(* IEC 61131-3 sources: iecf/tools/bench, 28 files *)

(* ---- fbcalls.st ---- *)
(* iecf's benchmark (docs/testing/performance.md): 10 instances of a FUNCTION_BLOCK and a FUNCTION called 50 times a cycle, a CTU.
   Standard IEC 61131-3, for both compilers: tools/bench/run.sh. *)
FUNCTION_BLOCK Filter
  VAR_INPUT x : DINT; k : DINT; END_VAR
  VAR_OUTPUT y : DINT; END_VAR
  VAR state : DINT; n : DINT; END_VAR
  state := state + (x - state) / k;
  n := n + 1;
  y := state + n MOD 7;
END_FUNCTION_BLOCK
FUNCTION Mix : DINT
  VAR_INPUT a : DINT; b : DINT; END_VAR
  Mix := (a * 3 + b) MOD 100003;
END_FUNCTION
PROGRAM main
  VAR f1 : Filter; f2 : Filter; f3 : Filter; f4 : Filter; f5 : Filter; f6 : Filter; f7 : Filter; f8 : Filter; f9 : Filter; f10 : Filter; c : CTU; i : INT; rep : INT; acc : DINT; END_VAR
  VAR o1 AT %QD0 : DINT; o2 AT %QW4 : INT; END_VAR
  FOR rep := 1 TO 50 DO
    FOR i := 1 TO 10 DO
      f1(x := acc + 1, k := 4);
      acc := Mix(a := acc, b := f1.y);
      f2(x := acc + 2, k := 4);
      acc := Mix(a := acc, b := f2.y);
      f3(x := acc + 3, k := 4);
      acc := Mix(a := acc, b := f3.y);
      f4(x := acc + 4, k := 4);
      acc := Mix(a := acc, b := f4.y);
      f5(x := acc + 5, k := 4);
      acc := Mix(a := acc, b := f5.y);
      f6(x := acc + 6, k := 4);
      acc := Mix(a := acc, b := f6.y);
      f7(x := acc + 7, k := 4);
      acc := Mix(a := acc, b := f7.y);
      f8(x := acc + 8, k := 4);
      acc := Mix(a := acc, b := f8.y);
      f9(x := acc + 9, k := 4);
      acc := Mix(a := acc, b := f9.y);
      f10(x := acc + 10, k := 4);
      acc := Mix(a := acc, b := f10.y);
    END_FOR;
    c(CU := NOT c.CU, PV := 30000);
  END_FOR;
  IF c.Q THEN c(R := TRUE); c(R := FALSE); END_IF;
  o1 := acc;
  o2 := c.CV;
END_PROGRAM
CONFIGURATION cf
  RESOURCE r ON x
    TASK tk(INTERVAL := T#10ms, PRIORITY := 1);
    PROGRAM p WITH tk : main;
  END_RESOURCE
END_CONFIGURATION

(* ---- m_fbcall.st ---- *)
(* iecf's benchmark (docs/testing/performance.md): a FUNCTION_BLOCK call.
   Standard IEC 61131-3, for both compilers: tools/bench/run.sh. *)
FUNCTION_BLOCK Acc
  VAR_INPUT x : DINT; k : DINT; END_VAR
  VAR_OUTPUT y : DINT; END_VAR
  y := (y + x * k) MOD 100000;
END_FUNCTION_BLOCK
PROGRAM main
  VAR i : DINT; f : Acc; n : DINT; END_VAR
  VAR o1 AT %QD0 : DINT; END_VAR
  FOR i := 1 TO 20000 DO
    f(x := i MOD 9, k := 2); n := f.y;
  END_FOR;
  o1 := n;
END_PROGRAM
CONFIGURATION cf
  RESOURCE r ON x
    TASK tk(INTERVAL := T#10ms, PRIORITY := 1);
    PROGRAM p WITH tk : main;
  END_RESOURCE
END_CONFIGURATION

(* ---- oo.st ---- *)
(* iecf's benchmark (docs/testing/performance.md): CODESYS's object
   orientation, iecf alone (--extension codesys): set `mode` to 0 for a
   method of an instance, 1 through an interface, 2 through a REFERENCE
   TO, 3 through a POINTER TO, 4 a property read through an interface. *)
INTERFACE ICounter
  METHOD Bump : DINT
    VAR_INPUT amount : DINT; END_VAR
  END_METHOD
  PROPERTY Value : DINT
  GET
  END_GET
  END_PROPERTY
END_INTERFACE
FUNCTION_BLOCK Base IMPLEMENTS ICounter
  VAR n : DINT; END_VAR
  METHOD PUBLIC Bump : DINT
    VAR_INPUT amount : DINT; END_VAR
    n := (n + amount) MOD 100003;
    Bump := n;
  END_METHOD
  PROPERTY PUBLIC Value : DINT
  GET
    Value := n;
  END_GET
  END_PROPERTY
END_FUNCTION_BLOCK
FUNCTION_BLOCK Derived EXTENDS Base
  METHOD PUBLIC Bump : DINT
    VAR_INPUT amount : DINT; END_VAR
    n := (n + amount * 2) MOD 100003;
    Bump := n;
  END_METHOD
END_FUNCTION_BLOCK
PROGRAM main
  VAR i : DINT; b : Base; d : Derived; c : ICounter; r : REFERENCE TO Base; p : POINTER TO Base;
      acc : DINT; mode : DINT; END_VAR
  VAR o1 AT %QD0 : DINT; END_VAR
  r REF= d;
  p := ADR(b);
  FOR i := 1 TO 20000 DO
    CASE mode OF
      0: acc := acc + b.Bump(amount := i MOD 7);
      1: c := d; acc := acc + c.Bump(amount := i MOD 7);
      2: acc := acc + r.Bump(amount := i MOD 7);
      3: acc := acc + p^.Bump(amount := i MOD 7);
      4: c := b; acc := acc + c.Value;
    END_CASE;
    acc := acc MOD 1000003;
  END_FOR;
  o1 := acc;
END_PROGRAM
CONFIGURATION cf
  RESOURCE r ON x
    TASK tk(INTERVAL := T#10ms, PRIORITY := 1);
    PROGRAM p WITH tk : main;
  END_RESOURCE
END_CONFIGURATION

(* ---- sfc.st ---- *)
(* iecf's benchmark (docs/testing/performance.md): 40 instances of a FUNCTION_BLOCK whose body is a four-step SFC chart of N actions.
   Standard IEC 61131-3, for both compilers: tools/bench/run.sh. *)
FUNCTION_BLOCK Machine
  VAR_INPUT seed : DINT; END_VAR
  VAR_OUTPUT work : DINT; cycles : DINT; END_VAR
  VAR n : DINT; acc : DINT; END_VAR
  INITIAL_STEP idle : start(N); END_STEP
  TRANSITION FROM idle TO fill := n >= 2; END_TRANSITION
  STEP fill : filling(N); END_STEP
  TRANSITION FROM fill TO heat := n >= 5; END_TRANSITION
  STEP heat : heating(N); END_STEP
  TRANSITION FROM heat TO drain := n >= 9; END_TRANSITION
  STEP drain : draining(N); END_STEP
  TRANSITION FROM drain TO idle := n >= 12; END_TRANSITION
  ACTION start :
    n := n + 1;
    acc := (acc * 7 + seed) MOD 100003;
    work := acc;
  END_ACTION
  ACTION filling :
    n := n + 1;
    acc := (acc + seed * 3) MOD 100003;
    work := acc;
  END_ACTION
  ACTION heating :
    n := n + 1;
    acc := (acc * 3 + 11) MOD 100003;
    work := acc;
  END_ACTION
  ACTION draining :
    n := n + 1;
    IF n >= 12 THEN n := 0; cycles := cycles + 1; END_IF;
    acc := (acc + 5) MOD 100003;
    work := acc;
  END_ACTION
END_FUNCTION_BLOCK
PROGRAM main
  VAR m1 : Machine; m2 : Machine; m3 : Machine; m4 : Machine; m5 : Machine; m6 : Machine; m7 : Machine; m8 : Machine; m9 : Machine; m10 : Machine; m11 : Machine; m12 : Machine; m13 : Machine; m14 : Machine; m15 : Machine; m16 : Machine; m17 : Machine; m18 : Machine; m19 : Machine; m20 : Machine; m21 : Machine; m22 : Machine; m23 : Machine; m24 : Machine; m25 : Machine; m26 : Machine; m27 : Machine; m28 : Machine; m29 : Machine; m30 : Machine; m31 : Machine; m32 : Machine; m33 : Machine; m34 : Machine; m35 : Machine; m36 : Machine; m37 : Machine; m38 : Machine; m39 : Machine; m40 : Machine; total : DINT; c : DINT; END_VAR
  VAR o1 AT %QD0 : DINT; o2 AT %QD4 : DINT; END_VAR
  total := 0; c := 0;
  m1(seed := 1); total := (total + m1.work) MOD 1000003; c := c + m1.cycles;
  m2(seed := 2); total := (total + m2.work) MOD 1000003; c := c + m2.cycles;
  m3(seed := 3); total := (total + m3.work) MOD 1000003; c := c + m3.cycles;
  m4(seed := 4); total := (total + m4.work) MOD 1000003; c := c + m4.cycles;
  m5(seed := 5); total := (total + m5.work) MOD 1000003; c := c + m5.cycles;
  m6(seed := 6); total := (total + m6.work) MOD 1000003; c := c + m6.cycles;
  m7(seed := 7); total := (total + m7.work) MOD 1000003; c := c + m7.cycles;
  m8(seed := 8); total := (total + m8.work) MOD 1000003; c := c + m8.cycles;
  m9(seed := 9); total := (total + m9.work) MOD 1000003; c := c + m9.cycles;
  m10(seed := 10); total := (total + m10.work) MOD 1000003; c := c + m10.cycles;
  m11(seed := 11); total := (total + m11.work) MOD 1000003; c := c + m11.cycles;
  m12(seed := 12); total := (total + m12.work) MOD 1000003; c := c + m12.cycles;
  m13(seed := 13); total := (total + m13.work) MOD 1000003; c := c + m13.cycles;
  m14(seed := 14); total := (total + m14.work) MOD 1000003; c := c + m14.cycles;
  m15(seed := 15); total := (total + m15.work) MOD 1000003; c := c + m15.cycles;
  m16(seed := 16); total := (total + m16.work) MOD 1000003; c := c + m16.cycles;
  m17(seed := 17); total := (total + m17.work) MOD 1000003; c := c + m17.cycles;
  m18(seed := 18); total := (total + m18.work) MOD 1000003; c := c + m18.cycles;
  m19(seed := 19); total := (total + m19.work) MOD 1000003; c := c + m19.cycles;
  m20(seed := 20); total := (total + m20.work) MOD 1000003; c := c + m20.cycles;
  m21(seed := 21); total := (total + m21.work) MOD 1000003; c := c + m21.cycles;
  m22(seed := 22); total := (total + m22.work) MOD 1000003; c := c + m22.cycles;
  m23(seed := 23); total := (total + m23.work) MOD 1000003; c := c + m23.cycles;
  m24(seed := 24); total := (total + m24.work) MOD 1000003; c := c + m24.cycles;
  m25(seed := 25); total := (total + m25.work) MOD 1000003; c := c + m25.cycles;
  m26(seed := 26); total := (total + m26.work) MOD 1000003; c := c + m26.cycles;
  m27(seed := 27); total := (total + m27.work) MOD 1000003; c := c + m27.cycles;
  m28(seed := 28); total := (total + m28.work) MOD 1000003; c := c + m28.cycles;
  m29(seed := 29); total := (total + m29.work) MOD 1000003; c := c + m29.cycles;
  m30(seed := 30); total := (total + m30.work) MOD 1000003; c := c + m30.cycles;
  m31(seed := 31); total := (total + m31.work) MOD 1000003; c := c + m31.cycles;
  m32(seed := 32); total := (total + m32.work) MOD 1000003; c := c + m32.cycles;
  m33(seed := 33); total := (total + m33.work) MOD 1000003; c := c + m33.cycles;
  m34(seed := 34); total := (total + m34.work) MOD 1000003; c := c + m34.cycles;
  m35(seed := 35); total := (total + m35.work) MOD 1000003; c := c + m35.cycles;
  m36(seed := 36); total := (total + m36.work) MOD 1000003; c := c + m36.cycles;
  m37(seed := 37); total := (total + m37.work) MOD 1000003; c := c + m37.cycles;
  m38(seed := 38); total := (total + m38.work) MOD 1000003; c := c + m38.cycles;
  m39(seed := 39); total := (total + m39.work) MOD 1000003; c := c + m39.cycles;
  m40(seed := 40); total := (total + m40.work) MOD 1000003; c := c + m40.cycles;
  o1 := total;
  o2 := c;
END_PROGRAM
CONFIGURATION cf
  RESOURCE r ON x
    TASK tk(INTERVAL := T#10ms, PRIORITY := 1);
    PROGRAM p WITH tk : main;
  END_RESOURCE
END_CONFIGURATION

(* ---- arith.st ---- *)
(* iecf's benchmark (docs/testing/performance.md): integer and LREAL arithmetic in a loop: DINT products and MOD, ROL and XOR of a DWORD, SQRT.
   Standard IEC 61131-3, for both compilers: tools/bench/run.sh. *)
PROGRAM main
  VAR i : DINT; acc : DINT; w : DWORD := 16#1234567; x : LREAL; END_VAR
  VAR o1 AT %QD0 : DINT; o2 AT %QD4 : DINT; o3 AT %QD8 : DWORD; END_VAR
  FOR i := 1 TO 20000 DO
    acc := (acc * 31 + i) MOD 1000003;
    w := ROL(w, 3) XOR DINT_TO_DWORD(i);
    x := x + SQRT(DINT_TO_LREAL(i)) * 0.5;
  END_FOR;
  IF x > 1.0E9 THEN x := 0.0; END_IF;
  o1 := acc;
  o2 := LREAL_TO_DINT(x);
  o3 := w;
END_PROGRAM
CONFIGURATION cf
  RESOURCE r ON x
    TASK tk(INTERVAL := T#10ms, PRIORITY := 1);
    PROGRAM p WITH tk : main;
  END_RESOURCE
END_CONFIGURATION

(* ---- m_bool.st ---- *)
(* iecf's benchmark (docs/testing/performance.md): BOOL logic and IF.
   Standard IEC 61131-3, for both compilers: tools/bench/run.sh. *)

PROGRAM main
  VAR i : DINT; b : BOOL; c : BOOL; n : DINT; END_VAR
  VAR o1 AT %QD0 : DINT; END_VAR
  FOR i := 1 TO 20000 DO
    b := (i MOD 3 = 0) XOR c; IF b AND NOT c THEN n := n + 1; END_IF; c := b OR (i MOD 5 = 1);
  END_FOR;
  o1 := n;
END_PROGRAM
CONFIGURATION cf
  RESOURCE r ON x
    TASK tk(INTERVAL := T#10ms, PRIORITY := 1);
    PROGRAM p WITH tk : main;
  END_RESOURCE
END_CONFIGURATION

(* ---- m_case.st ---- *)
(* iecf's benchmark (docs/testing/performance.md): CASE with lists and ranges.
   Standard IEC 61131-3, for both compilers: tools/bench/run.sh. *)

PROGRAM main
  VAR i : DINT; n : DINT; END_VAR
  VAR o1 AT %QD0 : DINT; END_VAR
  FOR i := 1 TO 20000 DO
    CASE i MOD 8 OF 0: n := n + 1; 1, 2: n := n + 2; 3..5: n := n - 1; ELSE n := n + 3; END_CASE;
  END_FOR;
  o1 := n;
END_PROGRAM
CONFIGURATION cf
  RESOURCE r ON x
    TASK tk(INTERVAL := T#10ms, PRIORITY := 1);
    PROGRAM p WITH tk : main;
  END_RESOURCE
END_CONFIGURATION

(* ---- m_empty.st ---- *)
(* iecf's benchmark (docs/testing/performance.md): one statement: the cost of a cycle itself.
   Standard IEC 61131-3, for both compilers: tools/bench/run.sh. *)
PROGRAM main
  VAR n : DINT; END_VAR
  VAR o1 AT %QD0 : DINT; END_VAR
  n := n + 1;
  o1 := n;
END_PROGRAM
CONFIGURATION cf
  RESOURCE r ON x
    TASK tk(INTERVAL := T#10ms, PRIORITY := 1);
    PROGRAM p WITH tk : main;
  END_RESOURCE
END_CONFIGURATION

(* ---- m_fcall.st ---- *)
(* iecf's benchmark (docs/testing/performance.md): a FUNCTION call.
   Standard IEC 61131-3, for both compilers: tools/bench/run.sh. *)
FUNCTION Add3 : DINT
  VAR_INPUT a : DINT; b : DINT; c : DINT; END_VAR
  Add3 := a + b + c;
END_FUNCTION
PROGRAM main
  VAR i : DINT; n : DINT; END_VAR
  VAR o1 AT %QD0 : DINT; END_VAR
  FOR i := 1 TO 20000 DO
    n := Add3(a := n, b := i, c := 1) MOD 100000;
  END_FOR;
  o1 := n;
END_PROGRAM
CONFIGURATION cf
  RESOURCE r ON x
    TASK tk(INTERVAL := T#10ms, PRIORITY := 1);
    PROGRAM p WITH tk : main;
  END_RESOURCE
END_CONFIGURATION

(* ---- m_iadd.st ---- *)
(* iecf's benchmark (docs/testing/performance.md): a DINT sum.
   Standard IEC 61131-3, for both compilers: tools/bench/run.sh. *)

PROGRAM main
  VAR i : DINT; acc : DINT; END_VAR
  VAR o1 AT %QD0 : DINT; END_VAR
  FOR i := 1 TO 20000 DO
    acc := acc + i MOD 7;
  END_FOR;
  o1 := acc;
END_PROGRAM
CONFIGURATION cf
  RESOURCE r ON x
    TASK tk(INTERVAL := T#10ms, PRIORITY := 1);
    PROGRAM p WITH tk : main;
  END_RESOURCE
END_CONFIGURATION

(* ---- m_iarr.st ---- *)
(* iecf's benchmark (docs/testing/performance.md): a DINT array element updated.
   Standard IEC 61131-3, for both compilers: tools/bench/run.sh. *)

PROGRAM main
  VAR i : DINT; a : ARRAY[0..63] OF DINT; k : DINT; END_VAR
  VAR o1 AT %QD0 : DINT; END_VAR
  FOR i := 1 TO 20000 DO
    k := i MOD 64; a[k] := a[k] + i MOD 5;
  END_FOR;
  o1 := a[3];
END_PROGRAM
CONFIGURATION cf
  RESOURCE r ON x
    TASK tk(INTERVAL := T#10ms, PRIORITY := 1);
    PROGRAM p WITH tk : main;
  END_RESOURCE
END_CONFIGURATION

(* ---- m_imul.st ---- *)
(* iecf's benchmark (docs/testing/performance.md): a DINT product and MOD.
   Standard IEC 61131-3, for both compilers: tools/bench/run.sh. *)

PROGRAM main
  VAR i : DINT; acc : DINT := 1; END_VAR
  VAR o1 AT %QD0 : DINT; END_VAR
  FOR i := 1 TO 20000 DO
    acc := (acc * 3 + i) MOD 65521;
  END_FOR;
  o1 := acc;
END_PROGRAM
CONFIGURATION cf
  RESOURCE r ON x
    TASK tk(INTERVAL := T#10ms, PRIORITY := 1);
    PROGRAM p WITH tk : main;
  END_RESOURCE
END_CONFIGURATION

(* ---- m_lradd.st ---- *)
(* iecf's benchmark (docs/testing/performance.md): an LREAL sum.
   Standard IEC 61131-3, for both compilers: tools/bench/run.sh. *)

PROGRAM main
  VAR i : DINT; x : LREAL; s : LREAL; END_VAR
  VAR o1 AT %QD0 : DINT; END_VAR
  FOR i := 1 TO 20000 DO
    x := DINT_TO_LREAL(i); s := s + x;
  END_FOR;
  o1 := LREAL_TO_DINT(s / 1000.0);
END_PROGRAM
CONFIGURATION cf
  RESOURCE r ON x
    TASK tk(INTERVAL := T#10ms, PRIORITY := 1);
    PROGRAM p WITH tk : main;
  END_RESOURCE
END_CONFIGURATION

(* ---- m_str.st ---- *)
(* iecf's benchmark (docs/testing/performance.md): CONCAT and LEN.
   Standard IEC 61131-3, for both compilers: tools/bench/run.sh. *)

PROGRAM main
  VAR i : DINT; s : STRING; n : DINT; END_VAR
  VAR o1 AT %QD0 : DINT; END_VAR
  FOR i := 1 TO 20000 DO
    s := CONCAT('ab', 'cd'); n := n + LEN(s);
  END_FOR;
  o1 := n;
END_PROGRAM
CONFIGURATION cf
  RESOURCE r ON x
    TASK tk(INTERVAL := T#10ms, PRIORITY := 1);
    PROGRAM p WITH tk : main;
  END_RESOURCE
END_CONFIGURATION

(* ---- m_struct.st ---- *)
(* iecf's benchmark (docs/testing/performance.md): a structure assigned field by field and copied.
   Standard IEC 61131-3, for both compilers: tools/bench/run.sh. *)
TYPE Pt : STRUCT x : DINT; y : DINT; END_STRUCT; END_TYPE
PROGRAM main
  VAR i : DINT; p : Pt; q : Pt; n : DINT; END_VAR
  VAR o1 AT %QD0 : DINT; END_VAR
  FOR i := 1 TO 20000 DO
    p.x := i; p.y := i MOD 9; q := p; n := (n + q.x + q.y) MOD 100000;
  END_FOR;
  o1 := n;
END_PROGRAM
CONFIGURATION cf
  RESOURCE r ON x
    TASK tk(INTERVAL := T#10ms, PRIORITY := 1);
    PROGRAM p WITH tk : main;
  END_RESOURCE
END_CONFIGURATION

(* ---- m_ton.st ---- *)
(* iecf's benchmark (docs/testing/performance.md): a TON called.
   Standard IEC 61131-3, for both compilers: tools/bench/run.sh. *)

PROGRAM main
  VAR i : DINT; t : TON; n : DINT; END_VAR
  VAR o1 AT %QD0 : DINT; END_VAR
  FOR i := 1 TO 20000 DO
    t(IN := i MOD 2 = 0, PT := T#5ms); IF t.Q THEN n := n + 1; END_IF;
  END_FOR;
  o1 := n;
END_PROGRAM
CONFIGURATION cf
  RESOURCE r ON x
    TASK tk(INTERVAL := T#10ms, PRIORITY := 1);
    PROGRAM p WITH tk : main;
  END_RESOURCE
END_CONFIGURATION

(* ---- m_while.st ---- *)
(* iecf's benchmark (docs/testing/performance.md): a WHILE loop.
   Standard IEC 61131-3, for both compilers: tools/bench/run.sh. *)

PROGRAM main
  VAR i : DINT; j : DINT; n : DINT; END_VAR
  VAR o1 AT %QD0 : DINT; END_VAR
  FOR i := 1 TO 20000 DO
    j := i MOD 8; WHILE j > 0 DO n := n + j; j := j - 1; END_WHILE;
  END_FOR;
  o1 := n;
END_PROGRAM
CONFIGURATION cf
  RESOURCE r ON x
    TASK tk(INTERVAL := T#10ms, PRIORITY := 1);
    PROGRAM p WITH tk : main;
  END_RESOURCE
END_CONFIGURATION

(* ---- r_arr.st ---- *)
(* iecf's benchmark (docs/testing/performance.md): a REAL array element updated through a computed index.
   Standard IEC 61131-3, for both compilers: tools/bench/run.sh. *)
PROGRAM main
  VAR i : DINT; k : INT; x : LREAL; s : LREAL; r : REAL; arr : ARRAY[1..64] OF REAL; END_VAR
  VAR o1 AT %QD0 : DINT; o2 AT %QD4 : DINT; o3 AT %QD8 : DINT; END_VAR
  FOR i := 1 TO 5000 DO
    x := DINT_TO_LREAL(i) * 0.001;
    k := DINT_TO_INT(i MOD 64) + 1; arr[k] := arr[k] * 0.5 + r / 1000.0; r := r + 0.25;
  END_FOR;
  IF s > 1.0E9 THEN s := 0.0; END_IF;
  o1 := LREAL_TO_DINT(s);
  o2 := REAL_TO_DINT(r);
  o3 := REAL_TO_DINT(arr[7] * 100.0);
END_PROGRAM
CONFIGURATION cf
  RESOURCE r ON x
    TASK tk(INTERVAL := T#10ms, PRIORITY := 1);
    PROGRAM p WITH tk : main;
  END_RESOURCE
END_CONFIGURATION

(* ---- r_conv.st ---- *)
(* iecf's benchmark (docs/testing/performance.md): one statement each: an LREAL product of a DINT, an LREAL sum.
   Standard IEC 61131-3, for both compilers: tools/bench/run.sh. *)
PROGRAM main
  VAR i : DINT; k : INT; x : LREAL; s : LREAL; r : REAL; arr : ARRAY[1..64] OF REAL; END_VAR
  VAR o1 AT %QD0 : DINT; o2 AT %QD4 : DINT; o3 AT %QD8 : DINT; END_VAR
  FOR i := 1 TO 5000 DO
    x := DINT_TO_LREAL(i) * 0.001;
    s := s + x;
  END_FOR;
  IF s > 1.0E9 THEN s := 0.0; END_IF;
  o1 := LREAL_TO_DINT(s);
  o2 := REAL_TO_DINT(r);
  o3 := REAL_TO_DINT(arr[7] * 100.0);
END_PROGRAM
CONFIGURATION cf
  RESOURCE r ON x
    TASK tk(INTERVAL := T#10ms, PRIORITY := 1);
    PROGRAM p WITH tk : main;
  END_RESOURCE
END_CONFIGURATION

(* ---- r_explog.st ---- *)
(* iecf's benchmark (docs/testing/performance.md): EXP of a negated variable plus LN.
   Standard IEC 61131-3, for both compilers: tools/bench/run.sh. *)
PROGRAM main
  VAR i : DINT; k : INT; x : LREAL; s : LREAL; r : REAL; arr : ARRAY[1..64] OF REAL; END_VAR
  VAR o1 AT %QD0 : DINT; o2 AT %QD4 : DINT; o3 AT %QD8 : DINT; END_VAR
  FOR i := 1 TO 5000 DO
    x := DINT_TO_LREAL(i) * 0.001;
    s := s + EXP(-x) + LN(1.0 + x);
  END_FOR;
  IF s > 1.0E9 THEN s := 0.0; END_IF;
  o1 := LREAL_TO_DINT(s);
  o2 := REAL_TO_DINT(r);
  o3 := REAL_TO_DINT(arr[7] * 100.0);
END_PROGRAM
CONFIGURATION cf
  RESOURCE r ON x
    TASK tk(INTERVAL := T#10ms, PRIORITY := 1);
    PROGRAM p WITH tk : main;
  END_RESOURCE
END_CONFIGURATION

(* ---- r_real.st ---- *)
(* iecf's benchmark (docs/testing/performance.md): a REAL product plus an LREAL converted.
   Standard IEC 61131-3, for both compilers: tools/bench/run.sh. *)
PROGRAM main
  VAR i : DINT; k : INT; x : LREAL; s : LREAL; r : REAL; arr : ARRAY[1..64] OF REAL; END_VAR
  VAR o1 AT %QD0 : DINT; o2 AT %QD4 : DINT; o3 AT %QD8 : DINT; END_VAR
  FOR i := 1 TO 5000 DO
    x := DINT_TO_LREAL(i) * 0.001;
    r := r * 0.999 + LREAL_TO_REAL(x);
  END_FOR;
  IF s > 1.0E9 THEN s := 0.0; END_IF;
  o1 := LREAL_TO_DINT(s);
  o2 := REAL_TO_DINT(r);
  o3 := REAL_TO_DINT(arr[7] * 100.0);
END_PROGRAM
CONFIGURATION cf
  RESOURCE r ON x
    TASK tk(INTERVAL := T#10ms, PRIORITY := 1);
    PROGRAM p WITH tk : main;
  END_RESOURCE
END_CONFIGURATION

(* ---- r_sincos.st ---- *)
(* iecf's benchmark (docs/testing/performance.md): SIN times COS.
   Standard IEC 61131-3, for both compilers: tools/bench/run.sh. *)
PROGRAM main
  VAR i : DINT; k : INT; x : LREAL; s : LREAL; r : REAL; arr : ARRAY[1..64] OF REAL; END_VAR
  VAR o1 AT %QD0 : DINT; o2 AT %QD4 : DINT; o3 AT %QD8 : DINT; END_VAR
  FOR i := 1 TO 5000 DO
    x := DINT_TO_LREAL(i) * 0.001;
    s := s + SIN(x) * COS(x);
  END_FOR;
  IF s > 1.0E9 THEN s := 0.0; END_IF;
  o1 := LREAL_TO_DINT(s);
  o2 := REAL_TO_DINT(r);
  o3 := REAL_TO_DINT(arr[7] * 100.0);
END_PROGRAM
CONFIGURATION cf
  RESOURCE r ON x
    TASK tk(INTERVAL := T#10ms, PRIORITY := 1);
    PROGRAM p WITH tk : main;
  END_RESOURCE
END_CONFIGURATION

(* ---- r_sqrtdiv.st ---- *)
(* iecf's benchmark (docs/testing/performance.md): SQRT divided by a sum.
   Standard IEC 61131-3, for both compilers: tools/bench/run.sh. *)
PROGRAM main
  VAR i : DINT; k : INT; x : LREAL; s : LREAL; r : REAL; arr : ARRAY[1..64] OF REAL; END_VAR
  VAR o1 AT %QD0 : DINT; o2 AT %QD4 : DINT; o3 AT %QD8 : DINT; END_VAR
  FOR i := 1 TO 5000 DO
    x := DINT_TO_LREAL(i) * 0.001;
    s := s + SQRT(x) / (1.0 + x * x);
  END_FOR;
  IF s > 1.0E9 THEN s := 0.0; END_IF;
  o1 := LREAL_TO_DINT(s);
  o2 := REAL_TO_DINT(r);
  o3 := REAL_TO_DINT(arr[7] * 100.0);
END_PROGRAM
CONFIGURATION cf
  RESOURCE r ON x
    TASK tk(INTERVAL := T#10ms, PRIORITY := 1);
    PROGRAM p WITH tk : main;
  END_RESOURCE
END_CONFIGURATION

(* ---- reals.st ---- *)
(* iecf's benchmark (docs/testing/performance.md): LREAL SIN, COS, EXP, LN, SQRT and a division, a REAL array, 5000 times a cycle.
   Standard IEC 61131-3, for both compilers: tools/bench/run.sh. *)
PROGRAM main
  VAR i : DINT; k : INT; x : LREAL; s : LREAL; r : REAL; arr : ARRAY[1..64] OF REAL; END_VAR
  VAR o1 AT %QD0 : DINT; o2 AT %QD4 : DINT; o3 AT %QD8 : DINT; END_VAR
  FOR i := 1 TO 5000 DO
    x := DINT_TO_LREAL(i) * 0.001;
    s := s + SIN(x) * COS(x) + EXP(-x) + LN(1.0 + x) + SQRT(x) / (1.0 + x * x);
    r := r * 0.999 + LREAL_TO_REAL(x);
    k := DINT_TO_INT(i MOD 64) + 1;
    arr[k] := arr[k] * 0.5 + r / 1000.0;
  END_FOR;
  IF s > 1.0E9 THEN s := 0.0; END_IF;
  o1 := LREAL_TO_DINT(s);
  o2 := REAL_TO_DINT(r);
  o3 := REAL_TO_DINT(arr[7] * 100.0);
END_PROGRAM
CONFIGURATION cf
  RESOURCE r ON x
    TASK tk(INTERVAL := T#10ms, PRIORITY := 1);
    PROGRAM p WITH tk : main;
  END_RESOURCE
END_CONFIGURATION

(* ---- realsf.st ---- *)
(* iecf's benchmark (docs/testing/performance.md): `reals` in REAL - SIN, COS, EXP, LN, SQRT and a division, a REAL array, 5000 times a cycle.
   Standard IEC 61131-3, for both compilers: tools/bench/run.sh. *)
PROGRAM main
  VAR i : DINT; k : INT; x : REAL; s : REAL; r : REAL; arr : ARRAY[1..64] OF REAL; END_VAR
  VAR o1 AT %QD0 : DINT; o2 AT %QD4 : DINT; o3 AT %QD8 : DINT; END_VAR
  FOR i := 1 TO 5000 DO
    x := DINT_TO_REAL(i) * 0.001;
    s := s + SIN(x) * COS(x) + EXP(-x) + LN(1.0 + x) + SQRT(x) / (1.0 + x * x);
    r := r * 0.999 + x;
    k := DINT_TO_INT(i MOD 64) + 1;
    arr[k] := arr[k] * 0.5 + r / 1000.0;
  END_FOR;
  IF s > 1.0E9 THEN s := 0.0; END_IF;
  o1 := REAL_TO_DINT(s);
  o2 := REAL_TO_DINT(r);
  o3 := REAL_TO_DINT(arr[7] * 100.0);
END_PROGRAM
CONFIGURATION cf
  RESOURCE r ON x
    TASK tk(INTERVAL := T#10ms, PRIORITY := 1);
    PROGRAM p WITH tk : main;
  END_RESOURCE
END_CONFIGURATION

(* ---- sort.st ---- *)
(* iecf's benchmark (docs/testing/performance.md): an insertion sort of 300 DINTs, filled by a linear congruential generator.
   Standard IEC 61131-3, for both compilers: tools/bench/run.sh. *)
PROGRAM main
  VAR a : ARRAY[1..300] OF DINT; i : INT; j : INT; k : DINT; seed : DINT := 7; sum : DINT; END_VAR
  VAR o1 AT %QD0 : DINT; o2 AT %QD4 : DINT; END_VAR
  FOR i := 1 TO 300 DO
    seed := (seed * 1103 + 12345) MOD 65536;
    a[i] := seed;
  END_FOR;
  FOR i := 2 TO 300 DO
    k := a[i];
    j := i - 1;
    WHILE j >= 1 DO
      IF a[j] <= k THEN EXIT; END_IF;
      a[j + 1] := a[j];
      j := j - 1;
    END_WHILE;
    a[j + 1] := k;
  END_FOR;
  sum := 0;
  FOR i := 1 TO 300 DO sum := (sum + a[i] * INT_TO_DINT(i)) MOD 1000003; END_FOR;
  o1 := sum;
  o2 := a[150];
END_PROGRAM
CONFIGURATION cf
  RESOURCE r ON x
    TASK tk(INTERVAL := T#10ms, PRIORITY := 1);
    PROGRAM p WITH tk : main;
  END_RESOURCE
END_CONFIGURATION

(* ---- strings.st ---- *)
(* iecf's benchmark (docs/testing/performance.md): CONCAT, LEFT, RIGHT, LEN, FIND, INT_TO_STRING and STRING_TO_INT, 1000 times a cycle.
   Standard IEC 61131-3, for both compilers: tools/bench/run.sh. *)
PROGRAM main
  VAR i : INT; s : STRING; t : STRING := 'pump-station-'; n : DINT; END_VAR
  VAR o1 AT %QD0 : DINT; END_VAR
  FOR i := 1 TO 1000 DO
    s := CONCAT(LEFT(t, 5 + i MOD 8), INT_TO_STRING(i));
    n := (n + LEN(s) + FIND(s, '9') + INT_TO_DINT(STRING_TO_INT(RIGHT(s, 1)))) MOD 1000003;
    IF s = 'pump-sta123' THEN n := n + 1; END_IF;
  END_FOR;
  o1 := n;
END_PROGRAM
CONFIGURATION cf
  RESOURCE r ON x
    TASK tk(INTERVAL := T#10ms, PRIORITY := 1);
    PROGRAM p WITH tk : main;
  END_RESOURCE
END_CONFIGURATION

(* ---- structs.st ---- *)
(* iecf's benchmark (docs/testing/performance.md): an array of 200 nested structures filled, copied through a FUNCTION's VAR_IN_OUT and reversed.
   Standard IEC 61131-3, for both compilers: tools/bench/run.sh. *)
TYPE
  Point : STRUCT x : DINT; y : DINT; END_STRUCT;
  Seg : STRUCT a : Point; b : Point; len2 : DINT; tag : INT; END_STRUCT;
END_TYPE
FUNCTION Measure : DINT
  VAR_IN_OUT s : Seg; END_VAR
  VAR dx : DINT; dy : DINT; END_VAR
  dx := s.b.x - s.a.x;
  dy := s.b.y - s.a.y;
  s.len2 := dx * dx + dy * dy;
  Measure := s.len2;
END_FUNCTION
PROGRAM main
  VAR segs : ARRAY[1..200] OF Seg; tmp : Seg; i : INT; rep : INT; acc : DINT; seed : DINT := 1; d : DINT; END_VAR
  VAR o1 AT %QD0 : DINT; o2 AT %QD4 : DINT; END_VAR
  FOR rep := 1 TO 20 DO
  FOR i := 1 TO 200 DO
    seed := (seed * 1103 + 12345) MOD 65536;
    segs[i].a.x := seed MOD 1000;
    segs[i].a.y := seed / 1000;
    segs[i].b := segs[i].a;
    segs[i].b.x := segs[i].b.x + INT_TO_DINT(i);
    segs[i].tag := i;
    tmp := segs[i];
    d := Measure(s := tmp);
    segs[i] := tmp;
  END_FOR;
  FOR i := 1 TO 100 DO
    tmp := segs[i];
    segs[i] := segs[201 - i];
    segs[201 - i] := tmp;
  END_FOR;
  END_FOR;
  acc := 0;
  FOR i := 1 TO 200 DO
    acc := (acc + segs[i].len2 * INT_TO_DINT(segs[i].tag)) MOD 1000003;
  END_FOR;
  o1 := acc;
  o2 := segs[1].a.x + segs[200].b.y;
END_PROGRAM
CONFIGURATION cf
  RESOURCE r ON x
    TASK tk(INTERVAL := T#10ms, PRIORITY := 1);
    PROGRAM p WITH tk : main;
  END_RESOURCE
END_CONFIGURATION
